Fanuc KAREL source: KA00049.KL

PROGRAM KA00049
%NOLOCKGROUP
VAR
  SRC: POSITION
  DST: INTEGER
BEGIN
  DST = SRC
END KA00049
